Universal Robots PolyScope program: program_1.urp

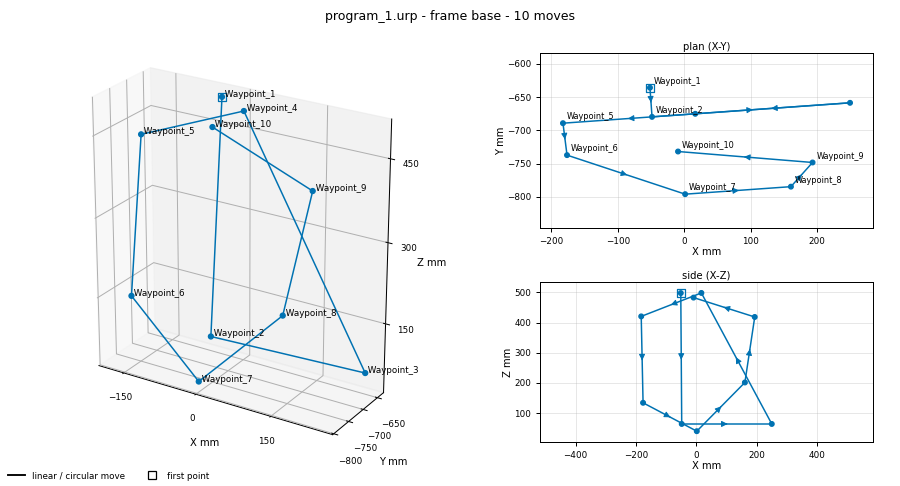
[picture p0: tool path of program_1.urp in frame base, 10 of 10 moves have a stored position in this frame; points joined in program order, loops and branches not executed]
Program program_1 (installation=default directory=/ursim/programs createdIn=3.15.8.106339 lastSavedIn=3.15.8.106339 robotSerialNumber=2018359999)
Calibrated DH parameters: a=[0, -0.425, -0.39225, 0, 0, 0]; d=[0.089159, 0, 0, 0.10915, 0.09465, 0.0823]; alpha=[1.570796, 0, 0, 1.570796, -1.570796, 0]; deltaTheta=[0, 0, 0, 0, 0, 0]
Robot Program (runOnlyOnce=false)
  Popup Message (haltProgram=false message=simulador letra L inputType=Text)
  MoveL speed 250 mm/s, acceleration 1200 mm/s^2 (useActiveTCP=true) feature=Base
    Waypoint Waypoint_1: TCP in base x=-51.679 y=-635.786 z=497.528 mm, rx=-0.0012 ry=3.1165 rz=0.0387 rad; joints [-84.997, -111.555, -54.056, -105.683, 91.544, 4.941] deg
    Waypoint Waypoint_2: TCP in base x=-48.565 y=-679.674 z=64.33 mm, rx=-0.0012 ry=3.1165 rz=0.0387 rad; joints [-85.058, -131.884, -89.022, -50.39, 91.543, 4.88] deg
    Waypoint Waypoint_3: TCP in base x=249.484 y=-658.527 z=64.33 mm, rx=-0.0012 ry=3.1165 rz=0.0387 rad; joints [-60.563, -134.278, -84.558, -51.704, 91.941, 29.383] deg
  Popup Message (haltProgram=false message=simulando letra o inputType=Text)
  MoveL speed 250 mm/s, acceleration 1200 mm/s^2 (useActiveTCP=true) feature=Base
    Waypoint Waypoint_4: TCP in base x=16.47 y=-675.06 z=497.928 mm, rx=-0.0012 ry=3.1165 rz=0.0387 rad; joints [-79.505, -118.01, -44.53, -108.599, 91.661, 10.433] deg
    Waypoint Waypoint_5: TCP in base x=-182.626 y=-689.186 z=420.33 mm, rx=-0.0012 ry=3.1165 rz=0.0387 rad; joints [-96.183, -121.822, -50.133, -99.614, 91.264, -6.245] deg
    Waypoint Waypoint_6: TCP in base x=-176.509 y=-737.272 z=134.333 mm, rx=-0.0012 ry=3.1165 rz=0.0387 rad; joints [-95.327, -135.559, -69.734, -66.256, 91.287, -5.389] deg
    Waypoint Waypoint_7: TCP in base x=1.295 y=-796.034 z=40.335 mm, rx=-0.0012 ry=3.1165 rz=0.0387 rad; joints [-82.193, -146.969, -63.048, -61.2, 91.605, 7.745] deg
    Waypoint Waypoint_8: TCP in base x=160.491 y=-784.738 z=201.601 mm, rx=-0.0012 ry=3.1165 rz=0.0387 rad; joints [-70.798, -138.395, -54.279, -78.202, 91.814, 19.144] deg
    Waypoint Waypoint_9: TCP in base x=193.064 y=-748.331 z=418.376 mm, rx=-0.0012 ry=3.1165 rz=0.0387 rad; joints [-67.614, -133.83, -30.47, -106.474, 91.86, 22.328] deg
    Waypoint Waypoint_10: TCP in base x=-9.411 y=-731.822 z=482.537 mm, rx=-0.0012 ry=3.1165 rz=0.0387 rad; joints [-82.342, -129.048, -28.851, -113.322, 91.602, 7.596] deg
